Fanuc KAREL source: KA00135.KL

PROGRAM KA00135
%NOLOCKGROUP
VAR
  SRC: ARRAY[2] OF SHORT
  DST: BOOLEAN
BEGIN
  SRC[1] = 2
  DST = SRC[1]
END KA00135
